{attribute 'qualified_only'}
VAR_GLOBAL
	
coffees 			: coffee;
teas				: tea;


END_VAR

(* stored: Version 1.1.0.1
   GVL gvl: Id {2a5719ea-eefe-42f9-8590-5791d8ba29d3} *)
